(* CODESYS project backup_pre_chaser_20261119.export

Project tree, tasks and I/O mapping:
  program PLC_PRG [ST]
  global variables GVL_IO
*)

// GVL_IO
VAR_GLOBAL
	xBtnStart AT %IX0.0 : BOOL;	// Nút START (UR20-8DI-P, kênh 0)
	xBtnStop  AT %IX0.1 : BOOL;	// Nút STOP (UR20-8DI-P, kênh 1)
	xBtnDir   AT %IX0.2 : BOOL;	// Nút ĐỔI CHIỀU chạy (UR20-8DI-P, kênh 2)
	byOut     AT %QB0   : BYTE;	// 8 ngõ ra UR20-8DO-P (bit 0..7 = kênh 0..7)
END_VAR

// PLC_PRG
PROGRAM PLC_PRG
VAR
	xRun      : BOOL;					// Đang chạy tuần tự
	xDirRev   : BOOL;					// FALSE: kênh 0 -> 7, TRUE: kênh 7 -> 0
	iStep     : INT := 0;				// Kênh đang sáng (0..7)
	tStepTime : TIME := T#500MS;		// Thời gian mỗi bước
	tStep     : TON;					// Timer bước
	rtStart   : R_TRIG;					// Sườn lên nút START
	rtStop    : R_TRIG;					// Sườn lên nút STOP
	rtDir     : R_TRIG;					// Sườn lên nút ĐỔI CHIỀU
END_VAR

// Phát hiện sườn lên của các nút nhấn
rtStart(CLK := GVL_IO.xBtnStart);
rtStop(CLK := GVL_IO.xBtnStop);
rtDir(CLK := GVL_IO.xBtnDir);

// START / STOP (STOP ưu tiên)
IF rtStop.Q THEN
	xRun := FALSE;
ELSIF rtStart.Q THEN
	xRun := TRUE;
END_IF

// Mỗi lần nhấn nút 3 thì đảo chiều chạy
IF rtDir.Q THEN
	xDirRev := NOT xDirRev;
END_IF

// Timer bước: tự reset sau mỗi chu kỳ
tStep(IN := xRun AND NOT tStep.Q, PT := tStepTime);

IF NOT xRun THEN
	iStep := 0;
	IF xDirRev THEN
		iStep := 7;
	END_IF
ELSIF tStep.Q THEN
	IF xDirRev THEN
		iStep := iStep - 1;
		IF iStep < 0 THEN
			iStep := 7;
		END_IF
	ELSE
		iStep := iStep + 1;
		IF iStep > 7 THEN
			iStep := 0;
		END_IF
	END_IF
END_IF

// Xuất ngõ ra: chỉ 1 kênh sáng tại mỗi thời điểm; STOP thì tắt hết
IF xRun THEN
	GVL_IO.byOut := SHL(BYTE#1, INT_TO_BYTE(iStep));
ELSE
	GVL_IO.byOut := 0;
END_IF

END_PROGRAM
